Fanuc KAREL source: kt00367.KL

-- PROVISIONAL review KL for V770-1; original PC SHA256 f6e4305d401f1cdbeb320fb0040f5f4e88806e38f12b9c68c54d560f259fe292
-- Incomplete behavior may be omitted. Consult companion uncertainty JSON. Do not deploy.
PROGRAM KT00367
%NOLOCKGROUP
VAR
  I1 : INTEGER
  OUT : BOOLEAN
-- UNRESOLVED_DECL Y2 type=002018
BEGIN
  -- UNRESOLVED_PC offsets 5-16; opcodes 2E,23
  -- UNRESOLVED_PC offsets 21-35; opcodes 2E,22,9D,33,B2
  -- UNRESOLVED_PC offsets 40-62; opcodes 21,22,9D,33,B1,5A,23
  -- UNRESOLVED_PC offsets 67-71; opcodes 7F
END KT00367
